(* IEC 61131-3 sources: codesys-framework/txt/application/ToDo/Hyperion, 15 files *)

(* ---- F_HyperionCreatePayloadString_1.pou.st ---- *)
FUNCTION F_HyperionCreatePayloadString_1 : ARRAY[0..63] OF BYTE
VAR_INPUT
	asEventPayload : ARRAY[1..10] OF STRING;
	iAmountPayload : INT;
END_VAR
VAR
	_sSeparator : STRING(1);
	_bySeparatorAsciiValue : BYTE;
	_byCharAsciiValue : BYTE;
	_iCounter : INT;
	_sPayloadPartString : STRING;
	_sPayloadString : STRING (cHYP_MAX_PAYLOADBYTESIZE);
	_iPayloadStringLength : INT;

	_abyPayloadByteArray : POINTER TO ARRAY [0 .. cHYP_MAX_PAYLOADBYTESIZE] OF BYTE;
	_abyPayloadByteArray_Return : ARRAY [0 .. cHYP_MAX_PAYLOADBYTESIZE] OF BYTE;
END_VAR

// --- BEGIN IMPLEMENTATION ---

// Init
_sPayloadString := '';
_sSeparator := ';';
_bySeparatorAsciiValue := 59;
// Check PayloadStrings
FOR _iCounter := 1 TO iAmountPayload BY 1 DO
	_sPayloadPartString := CONCAT(STR1 := asEventPayload[_iCounter], STR2 := _sSeparator);
	_sPayloadString := CONCAT(STR1 := _sPayloadString, STR2 := _sPayloadPartString);
END_FOR

// String to ByteArray
_iPayloadStringLength := LEN (STR := _sPayloadString);
_abyPayloadByteArray := ADR (_sPayloadString);

// Replace ';' with 0
FOR _iCounter := 0 TO cHYP_MAX_PAYLOADBYTESIZE BY 1 DO
	IF _iCounter < _iPayloadStringLength THEN
		_byCharAsciiValue := _abyPayloadByteArray^[_iCounter];
 		IF (_byCharAsciiValue <> _bySeparatorAsciiValue) THEN
			_abyPayloadByteArray_Return[_iCounter] := _byCharAsciiValue;
		ELSE
			_abyPayloadByteArray_Return[_iCounter] := 0;
		END_IF
	ELSE
		_abyPayloadByteArray_Return[_iCounter] := 0;
	END_IF
END_FOR

F_HyperionCreatePayloadString := _abyPayloadByteArray_Return;

(* ---- F_ParameterHandler_Bool.pou.st ---- *)
FUNCTION F_ParameterHandler_Bool : BOOL
VAR_INPUT
	eSubMachine 				: INT;
	w 							: WORD;
	eMode 						: E_ParameterMode;
	udiParameterId 				: UDINT;
	xExternalValidationFailed 	: BOOL := FALSE;
END_VAR
VAR_IN_OUT
	xValidationFailed 			: BOOL;
END_VAR
VAR_IN_OUT
	xHypValue 					: BOOL;
	xPLCValue 					: BOOL;
END_VAR
VAR
	_xParameterValid 			: BOOL;
	_rHypValue 					: REAL;
	_rPLCValue 					: REAL;
END_VAR

// --- BEGIN IMPLEMENTATION ---

IF (eMode = E_ParameterMode.Invalid) THEN
	xValidationFailed := TRUE;
	RETURN;
END_IF

IF xHypValue THEN
	_rHypValue := 1;
ELSE
	_rHypValue := 0;
END_IF

IF xPLCValue THEN
	_rPLCValue := 1;
ELSE
	_rPLCValue := 0;
END_IF

F_ParameterHandler_Real (
	eSubMachine := eSubMachine,
	w := w,
	eMode := eMode,
	udiParameterId := udiParameterId,
	xCanBeZero := TRUE,
	rLowLimit := 0,
	rUppLimit := 1,
	xValidationFailed := xValidationFailed,
	xExternalValidationFailed := xExternalValidationFailed,
	rHypValue := _rHypValue,
	rPLCValue := _rPLCValue);

xHypValue := _rHypValue = 1;
xPLCValue := _rPLCValue = 1;

(* ---- F_ParameterHandler_DInt.pou.st ---- *)
FUNCTION F_ParameterHandler_DInt : BOOL
VAR_INPUT
	eSubMachine 				: INT;
	w 							: WORD;
	eMode 						: E_ParameterMode;
	udiParameterId 				: UDINT;
	xCanBeZero 					: BOOL;
	diLowLimit 					: DINT;
	diUppLimit 					: DINT;
	xExternalValidationFailed 	: BOOL := FALSE;
END_VAR
VAR_IN_OUT
	xValidationFailed 			: BOOL;
	diHypValue 					: DINT;
	diPLCValue 					: DINT;
END_VAR
VAR
	_xParameterValid 			: BOOL;
	_rHypValue 					: REAL;
	_rPLCValue 					: REAL;
END_VAR

// --- BEGIN IMPLEMENTATION ---

IF eMode = E_ParameterMode.Invalid THEN
	xValidationFailed := TRUE;
	RETURN;
END_IF

_rHypValue := DINT_TO_REAL (diHypValue);
_rPLCValue := DINT_TO_REAL (diPLCValue);

F_ParameterHandler_Real (
	eSubMachine := eSubMachine,
	w := w,
	eMode := eMode,
	udiParameterId := udiParameterId,
	xCanBeZero := xCanBeZero,
	rLowLimit := DINT_TO_REAL (diLowLimit),
	rUppLimit := DINT_TO_REAL (diUppLimit),
	xValidationFailed := xValidationFailed,
	xExternalValidationFailed := xExternalValidationFailed,
	rHypValue := _rHypValue,
	rPLCValue := _rPLCValue);

diHypValue := REAL_TO_DINT (_rHypValue);
diPLCValue := REAL_TO_DINT (_rPLCValue);

(* ---- F_ParameterHandler_DWord.pou.st ---- *)
FUNCTION F_ParameterHandler_DWord : BOOL
VAR_INPUT
	eSubMachine 				: INT;
	w 							: WORD;
	eMode 						: E_ParameterMode;
	udiParameterId 				: UDINT;
	xCanBeZero 					: BOOL;
	dwLowLimit 					: DWORD;
	dwUppLimit 					: DWORD;
	xExternalValidationFailed 	: BOOL := FALSE;
END_VAR
VAR_IN_OUT
	xValidationFailed 			: BOOL;
	dwHypValue 					: DWORD;
	dwPLCValue 					: DWORD;
END_VAR
VAR
	_xParameterValid 			: BOOL;
	_rHypValue 					: REAL;
	_rPLCValue 					: REAL;
END_VAR

// --- BEGIN IMPLEMENTATION ---

IF eMode = E_ParameterMode.Invalid THEN
	xValidationFailed := TRUE;
	RETURN;
END_IF

_rHypValue := DWORD_TO_REAL (dwHypValue);
_rPLCValue := DWORD_TO_REAL (dwPLCValue);

F_ParameterHandler_Real (
	eSubMachine := eSubMachine,
	w := w,
	eMode := eMode,
	udiParameterId := udiParameterId,
	xCanBeZero := xCanBeZero,
	rLowLimit := DWORD_TO_REAL (dwLowLimit),
	rUppLimit := DWORD_TO_REAL (dwUppLimit),
	xValidationFailed := xValidationFailed,
	xExternalValidationFailed := xExternalValidationFailed,
	rHypValue := _rHypValue,
	rPLCValue := _rPLCValue);

dwHypValue := REAL_TO_DWORD (_rHypValue);
dwPLCValue := REAL_TO_DWORD (_rPLCValue);

(* ---- F_ParameterHandler_Int.pou.st ---- *)
FUNCTION F_ParameterHandler_Int : BOOL
VAR_INPUT
	eSubMachine 				: INT;
	w 							: WORD;
	eMode 						: E_ParameterMode;
	udiParameterId 				: UDINT;
	xCanBeZero 					: BOOL;
	iLowLimit 					: INT;
	iUppLimit 					: INT;
	xExternalValidationFailed 	: BOOL := FALSE;
END_VAR
VAR_IN_OUT
	xValidationFailed 			: BOOL;
	iHypValue 					: INT;
	iPLCValue 					: INT;
END_VAR
VAR
	_xParameterValid 			: BOOL;
	_rHypValue 					: REAL;
	_rPLCValue 					: REAL;
END_VAR

// --- BEGIN IMPLEMENTATION ---

IF eMode = E_ParameterMode.Invalid THEN
	xValidationFailed := TRUE;
	RETURN;
END_IF

_rHypValue := INT_TO_REAL (iHypValue);
_rPLCValue := INT_TO_REAL (iPLCValue);

F_ParameterHandler_Real (
	eSubMachine := eSubMachine,
	w := w,
	eMode := eMode,
	udiParameterId := udiParameterId,
	xCanBeZero := xCanBeZero,
	rLowLimit := INT_TO_REAL (iLowLimit),
	rUppLimit := INT_TO_REAL (iUppLimit),
	xValidationFailed := xValidationFailed,
	xExternalValidationFailed := xExternalValidationFailed,
	rHypValue := _rHypValue,
	rPLCValue := _rPLCValue);

iHypValue := REAL_TO_INT (_rHypValue);
iPLCValue := REAL_TO_INT (_rPLCValue);

(* ---- F_ParameterHandler_LReal.pou.st ---- *)
FUNCTION F_ParameterHandler_LReal : BOOL
VAR_INPUT
	eSubMachine 				: INT;
	w 							: WORD;
	eMode 						: E_ParameterMode;
	udiParameterId 				: UDINT;
	xCanBeZero 					: BOOL;
	lrLowLimit 					: LREAL;
	lrUppLimit 					: LREAL;
	xExternalValidationFailed 	: BOOL := FALSE;
END_VAR
VAR_IN_OUT
	xValidationFailed 			: BOOL;
	lrHypValue 					: LREAL;
	lrPLCValue 					: LREAL;
END_VAR
VAR
	_xParameterValid 			: BOOL;
END_VAR

// --- BEGIN IMPLEMENTATION ---

// Check
IF eMode = E_ParameterMode.Invalid THEN
	xValidationFailed := TRUE;
	RETURN;
END_IF

// Check HypValues
IF eMode = E_ParameterMode.CheckHyp THEN
	_xParameterValid := TRUE;
	IF NOT xCanBeZero AND lrHypValue = 0 THEN
		_xParameterValid := FALSE;
	ELSIF lrHypValue < lrLowLimit THEN
		_xParameterValid := FALSE;
	ELSIF lrHypValue > lrUppLimit THEN
		_xParameterValid := FALSE;
	ELSIF xExternalValidationFailed THEN
		_xParameterValid := FALSE;
	END_IF

	// !!!!! SET xParameterValidationFailed (Reset will be performed elsewhere)
	IF NOT _xParameterValid THEN
		xValidationFailed := TRUE;
	END_IF
END_IF

// Check PLCValues
IF eMode = E_ParameterMode.CheckPLC THEN
	_xParameterValid := TRUE;
	IF NOT xCanBeZero AND lrPLCValue = 0 THEN
		_xParameterValid := FALSE;
	ELSIF lrPLCValue < lrLowLimit THEN
		_xParameterValid := FALSE;
	ELSIF lrPLCValue > lrUppLimit THEN
		_xParameterValid := FALSE;
	ELSIF xExternalValidationFailed THEN
		_xParameterValid := FALSE;
	END_IF

	// !!!!! SET xParameterValidationFailed (Reset will be performed elsewhere)
	IF NOT _xParameterValid THEN
		xValidationFailed := TRUE;
	END_IF
END_IF

// Validate HyperionValues
IF eMode = E_ParameterMode.ValidateHyp OR eMode = E_ParameterMode.ValidateHypAndSavePLC THEN
	_xParameterValid := TRUE;
	IF NOT xCanBeZero AND lrHypValue = 0 THEN
		_xParameterValid := FALSE;
		// Insert message parametervalue is Zero
		F_Event_InsertMessage_ParameterChange (
			eSubMachine := eSubMachine,
			w := w,
			eValidationCode := E_ParameterValidationCode.Validation_Failed_IsZero,
			udiEventID := udiParameterId,
			rParameterValue_New := lrHypValue,
			rParameterValue_Previous := lrPLCValue,
			rParameterValue_MinimumValue := LREAL_TO_REAL(lrLowLimit),
			rParameterValue_MaximumValue := LREAL_TO_REAL(lrUppLimit));
	ELSIF lrHypValue < lrLowLimit THEN
		_xParameterValid := FALSE;
		//Insert message parametervalue < rValueLowerLimit
		F_Event_InsertMessage_ParameterChange (
			eSubMachine := eSubMachine,
			w := w,
			eValidationCode := E_ParameterValidationCode.Validation_Failed_BelowMinimum,
			udiEventID := udiParameterId,
			rParameterValue_New := lrHypValue,
			rParameterValue_Previous := lrPLCValue,
			rParameterValue_MinimumValue := LREAL_TO_REAL(lrLowLimit),
			rParameterValue_MaximumValue := LREAL_TO_REAL(lrUppLimit));
	ELSIF lrHypValue > lrUppLimit THEN
		_xParameterValid := FALSE;
		// Insert message parametervalue > rValueUpperLimit
		F_Event_InsertMessage_ParameterChange (
			eSubMachine := eSubMachine,
			w := w,
			eValidationCode := E_ParameterValidationCode.Validation_Failed_AboveMaximum,
			udiEventID := udiParameterId,
			rParameterValue_New := lrHypValue,
			rParameterValue_Previous := lrPLCValue,
			rParameterValue_MinimumValue := LREAL_TO_REAL(lrLowLimit),
			rParameterValue_MaximumValue := LREAL_TO_REAL(lrUppLimit));
	ELSIF xExternalValidationFailed THEN
		_xParameterValid := FALSE;
		// Insert message externalvalidationfailed
		F_Event_InsertMessage_ParameterChange (
			eSubMachine := eSubMachine,
			w := w,
			eValidationCode := E_ParameterValidationCode.Validation_Failed_External,
			udiEventID := udiParameterId,
			rParameterValue_New := lrHypValue,
			rParameterValue_Previous := lrPLCValue,
			rParameterValue_MinimumValue := LREAL_TO_REAL(lrLowLimit),
			rParameterValue_MaximumValue := LREAL_TO_REAL(lrUppLimit));
	END_IF

	// !!!!! SET xParameterValidationFailed (Reset will be performed elsewhere)
	IF NOT _xParameterValid THEN
		xValidationFailed := TRUE;
	END_IF
END_IF

// Save
IF eMode = E_ParameterMode.SavePLC OR (eMode = E_ParameterMode.ValidateHypAndSavePLC AND _xParameterValid) THEN
	IF lrPLCValue <> lrHypValue THEN
		F_Event_InsertMessage_ParameterChange (
			eSubMachine := eSubMachine,
			w := w,
			eValidationCode := E_ParameterValidationCode.Validation_Ok,
			udiEventID := udiParameterId,
			rParameterValue_New := lrHypValue,
			rParameterValue_Previous := lrPLCValue,
			rParameterValue_MinimumValue := LREAL_TO_REAL(lrLowLimit),
			rParameterValue_MaximumValue := LREAL_TO_REAL(lrUppLimit));
		lrPLCValue := lrHypValue;
	END_IF
END_IF

// Copy
IF eMode = E_ParameterMode.CopyPLCToHyp THEN
	lrHypValue := lrPLCValue;
END_IF

(* ---- F_ParameterHandler_Real.pou.st ---- *)
FUNCTION F_ParameterHandler_Real : BOOL
VAR_INPUT
	eSubMachine 				: INT;
	w 							: WORD;
	eMode 						: E_ParameterMode;
	udiParameterId 				: UDINT;
	xCanBeZero 					: BOOL;
	rLowLimit 					: REAL;
	rUppLimit 					: REAL;
	xExternalValidationFailed 	: BOOL := FALSE;
END_VAR
VAR_IN_OUT
	xValidationFailed 			: BOOL;
	rHypValue 					: REAL;
	rPLCValue 					: REAL;
END_VAR
VAR
	_xParameterValid 			: BOOL;
END_VAR

// --- BEGIN IMPLEMENTATION ---

// Check
IF eMode = E_ParameterMode.Invalid THEN
	xValidationFailed := TRUE;
	RETURN;
END_IF

// Check HypValues
IF eMode = E_ParameterMode.CheckHyp THEN
	_xParameterValid := TRUE;
	IF NOT xCanBeZero AND rHypValue = 0 THEN
		_xParameterValid := FALSE;
	ELSIF rHypValue < rLowLimit THEN
		_xParameterValid := FALSE;
	ELSIF rHypValue > rUppLimit THEN
		_xParameterValid := FALSE;
	ELSIF xExternalValidationFailed THEN
		_xParameterValid := FALSE;
	END_IF

	// !!!!! SET xParameterValidationFailed (Reset will be performed elsewhere)
	IF NOT _xParameterValid THEN
		xValidationFailed := TRUE;
	END_IF
END_IF

// Check PLCValues
IF eMode = E_ParameterMode.CheckPLC THEN
	_xParameterValid := TRUE;
	IF NOT xCanBeZero AND rPLCValue = 0 THEN
		_xParameterValid := FALSE;
	ELSIF rPLCValue < rLowLimit THEN
		_xParameterValid := FALSE;
	ELSIF rPLCValue > rUppLimit THEN
		_xParameterValid := FALSE;
	ELSIF xExternalValidationFailed THEN
		_xParameterValid := FALSE;
	END_IF

	// !!!!! SET xParameterValidationFailed (Reset will be performed elsewhere)
	IF NOT _xParameterValid THEN
		xValidationFailed := TRUE;
	END_IF
END_IF

// Validate HyperionValues
IF eMode = E_ParameterMode.ValidateHyp OR eMode = E_ParameterMode.ValidateHypAndSavePLC THEN
	_xParameterValid := TRUE;
	IF NOT xCanBeZero AND rHypValue = 0 THEN
		_xParameterValid := FALSE;
		// Insert message parametervalue is Zero
		F_Event_InsertMessage_ParameterChange (
			eSubMachine := eSubMachine,
			w := w,
			eValidationCode := E_ParameterValidationCode.Validation_Failed_IsZero,
			udiEventID := udiParameterId,
			rParameterValue_New := rHypValue,
			rParameterValue_Previous := rPLCValue,
			rParameterValue_MinimumValue := rLowLimit,
			rParameterValue_MaximumValue := rUppLimit);
	ELSIF rHypValue < rLowLimit THEN
		_xParameterValid := FALSE;
		//Insert message parametervalue < rValueLowerLimit
		F_Event_InsertMessage_ParameterChange (
			eSubMachine := eSubMachine,
			w := w,
			eValidationCode := E_ParameterValidationCode.Validation_Failed_BelowMinimum,
			udiEventID := udiParameterId,
			rParameterValue_New := rHypValue,
			rParameterValue_Previous := rPLCValue,
			rParameterValue_MinimumValue := rLowLimit,
			rParameterValue_MaximumValue := rUppLimit);
	ELSIF rHypValue > rUppLimit THEN
		_xParameterValid := FALSE;
		// Insert message parametervalue > rValueUpperLimit
		F_Event_InsertMessage_ParameterChange (
			eSubMachine := eSubMachine,
			w := w,
			eValidationCode := E_ParameterValidationCode.Validation_Failed_AboveMaximum,
			udiEventID := udiParameterId,
			rParameterValue_New := rHypValue,
			rParameterValue_Previous := rPLCValue,
			rParameterValue_MinimumValue := rLowLimit,
			rParameterValue_MaximumValue := rUppLimit);
	ELSIF xExternalValidationFailed THEN
		_xParameterValid := FALSE;
		// Insert message externalvalidationfailed
		F_Event_InsertMessage_ParameterChange (
			eSubMachine := eSubMachine,
			w := w,
			eValidationCode := E_ParameterValidationCode.Validation_Failed_External,
			udiEventID := udiParameterId,
			rParameterValue_New := rHypValue,
			rParameterValue_Previous := rPLCValue,
			rParameterValue_MinimumValue := rLowLimit,
			rParameterValue_MaximumValue := rUppLimit);
	END_IF

	// !!!!! SET xParameterValidationFailed (Reset will be performed elsewhere)
	IF NOT _xParameterValid THEN
		xValidationFailed := TRUE;
	END_IF
END_IF

// Save
IF eMode = E_ParameterMode.SavePLC OR (eMode = E_ParameterMode.ValidateHypAndSavePLC AND _xParameterValid) THEN
	IF rPLCValue <> rHypValue THEN
		F_Event_InsertMessage_ParameterChange (
			eSubMachine := eSubMachine,
			w := w,
			eValidationCode := E_ParameterValidationCode.Validation_Ok,
			udiEventID := udiParameterId,
			rParameterValue_New := rHypValue,
			rParameterValue_Previous := rPLCValue,
			rParameterValue_MinimumValue := rLowLimit,
			rParameterValue_MaximumValue := rUppLimit);
		rPLCValue := rHypValue;
	END_IF
END_IF

// Copy
IF eMode = E_ParameterMode.CopyPLCToHyp THEN
	rHypValue := rPLCValue;
END_IF

(* ---- F_ParameterHandler_String.pou.st ---- *)
FUNCTION F_ParameterHandler_String : BOOL
VAR_INPUT
	eSubMachine 				: INT;
	w 							: WORD;
	eMode 						: E_ParameterMode;
	udiParameterId 				: UDINT;
	xCanBeLengthZero 			: BOOL;
	iLowLengthLimit 			: INT;
	iUppLengthLimit 			: INT;
	xExternalValidationFailed 	: BOOL := FALSE;
END_VAR
VAR_IN_OUT
	xValidationFailed 			: BOOL;
	sHypValue 					: STRING;
	sPLCValue 					: STRING;
END_VAR
VAR
	_xParameterValid 			: BOOL;
	_sHypValue 					: STRING;
	_sPLCValue 					: STRING;
END_VAR

// --- BEGIN IMPLEMENTATION ---

_sHypValue := sHypValue;
_sPLCValue := sPLCValue;

// Check
IF (eMode = E_ParameterMode.Invalid) THEN
	xValidationFailed := TRUE;
	RETURN;
END_IF

// Check HypValues
IF (eMode = E_ParameterMode.CheckHyp) THEN
	_xParameterValid := TRUE;
	IF NOT xCanBeLengthZero AND (_sHypValue = '') THEN
		_xParameterValid := FALSE;
	ELSIF (LEN (_sHypValue) < iLowLengthLimit) THEN
		_xParameterValid := FALSE;
	ELSIF (LEN (_sHypValue) > iUppLengthLimit) THEN
		_xParameterValid := FALSE;
	ELSIF xExternalValidationFailed THEN
		_xParameterValid := FALSE;
	END_IF
	// !!!!!  SET xParameterValidationFailed (Reset will be performed elsewhere)
	IF (_xParameterValid = FALSE) THEN
		xValidationFailed := TRUE;
	END_IF
END_IF

//Check PLCValues
IF (eMode = E_ParameterMode.CheckPLC) THEN
	_xParameterValid := TRUE;
	IF (NOT xCanBeLengthZero AND (_sPLCValue = '')) THEN
		_xParameterValid := FALSE;
	ELSIF (LEN (_sPLCValue) < iLowLengthLimit) THEN
		_xParameterValid := FALSE;
	ELSIF (LEN (_sPLCValue) > iUppLengthLimit) THEN
		_xParameterValid := FALSE;
	ELSIF xExternalValidationFailed THEN
		_xParameterValid := FALSE;
	END_IF
	// !!!!!  SET xParameterValidationFailed (Reset will be performed elsewhere)
	IF NOT _xParameterValid THEN
		xValidationFailed := TRUE;
	END_IF
END_IF

// Validate HyperionValues
IF ((eMode = E_ParameterMode.ValidateHyp) OR (eMode = E_ParameterMode.ValidateHypAndSavePLC)) THEN
	_xParameterValid := TRUE;
	IF (NOT xCanBeLengthZero AND (_sHypValue = '')) THEN
		_xParameterValid := FALSE;
		// Insert message parametervalue is Zero
		F_Event_InsertMessage_StringParameterChange (
			eSubMachine := eSubMachine,
			w := w,
			udiEventID := udiParameterId,
			eValidationCode := E_ParameterValidationCode.Validation_Failed_IsZero,
			sParameterValue_Previous := _sPLCValue,
			sParameterValue_New := _sHypValue,
			iParameterValue_MinimumValue := iLowLengthLimit,
			iParameterValue_MaximumValue := iUppLengthLimit);
	ELSIF (LEN (_sHypValue) < iLowLengthLimit) THEN
		_xParameterValid := FALSE;
		// Insert message parametervalue < rValueLowerLimit
		F_Event_InsertMessage_StringParameterChange (
			eSubMachine := eSubMachine,
			w := w,
			udiEventID := udiParameterId,
			eValidationCode := E_ParameterValidationCode.Validation_Failed_BelowMinimum,
			sParameterValue_Previous := _sPLCValue,
			sParameterValue_New := _sHypValue,
			iParameterValue_MinimumValue := iLowLengthLimit,
			iParameterValue_MaximumValue := iUppLengthLimit);
	ELSIF (LEN (_sHypValue) > iUppLengthLimit) THEN
		_xParameterValid := FALSE;
		// Insert message parametervalue > rValueUpperLimit
		F_Event_InsertMessage_StringParameterChange (
			eSubMachine := eSubMachine,
			w := w,
			udiEventID := udiParameterId,
			eValidationCode := E_ParameterValidationCode.Validation_Failed_AboveMaximum,
			sParameterValue_Previous := _sPLCValue,
			sParameterValue_New := _sHypValue,
			iParameterValue_MinimumValue := iLowLengthLimit,
			iParameterValue_MaximumValue := iUppLengthLimit);
	ELSIF xExternalValidationFailed THEN
		_xParameterValid := FALSE;
		// Insert message external validatio nfailed
		F_Event_InsertMessage_StringParameterChange (
			eSubMachine := eSubMachine,
			w := w,
			udiEventID := udiParameterId,
			eValidationCode := E_ParameterValidationCode.Validation_Failed_External,
			sParameterValue_Previous := _sPLCValue,
			sParameterValue_New := _sHypValue,
			iParameterValue_MinimumValue := iLowLengthLimit,
			iParameterValue_MaximumValue := iUppLengthLimit);
	END_IF
	// !!!!!  SET xParameterValidationFailed (Reset will be performed elsewhere)
	IF NOT _xParameterValid THEN
		xValidationFailed := TRUE;
	END_IF
END_IF

// Save
IF ((eMode = E_ParameterMode.SavePLC) OR ((eMode = E_ParameterMode.ValidateHypAndSavePLC) AND _xParameterValid)) THEN
	IF (_sPLCValue <> _sHypValue) THEN
		F_Event_InsertMessage_StringParameterChange (
			eSubMachine := eSubMachine,
			w :=w,
			udiEventID := udiParameterId,
			eValidationCode := E_ParameterValidationCode.Validation_Ok,
			sParameterValue_Previous := _sPLCValue,
			sParameterValue_New := _sHypValue,
			iParameterValue_MinimumValue := iLowLengthLimit,
			iParameterValue_MaximumValue := iUppLengthLimit);
		_sPLCValue := _sHypValue;
	END_IF
END_IF

// Copy
IF (eMode = E_ParameterMode.CopyPLCToHyp) THEN
	_sHypValue := _sPLCValue;
END_IF

sHypValue := _sHypValue;
sPLCValue := _sPLCValue;

(* ---- F_ParameterHandler_UDInt.pou.st ---- *)
FUNCTION F_ParameterHandler_UDInt : BOOL
VAR_INPUT
	eSubMachine 				: INT;
	w 							: WORD;
	eMode 						: E_ParameterMode;
	udiParameterId	 			: UDINT;
	xCanBeZero 					: BOOL;
	udiLowLimit 				: UDINT;
	udiUppLimit 				: UDINT;
	xExternalValidationFailed 	: BOOL := FALSE;
END_VAR
VAR_IN_OUT
	xValidationFailed 			: BOOL;
	udiHypValue 				: UDINT;
	udiPLCValue 				: UDINT;
END_VAR
VAR
	_xParameterValid 			: BOOL;
	_rHypValue 					: REAL;
	_rPLCValue 					: REAL;
END_VAR

// --- BEGIN IMPLEMENTATION ---

IF eMode = E_ParameterMode.Invalid THEN
	xValidationFailed := TRUE;
	RETURN;
END_IF

_rHypValue := UDINT_TO_REAL (udiHypValue);
_rPLCValue := UDINT_TO_REAL (udiPLCValue);

F_ParameterHandler_Real (
	eSubMachine := eSubMachine,
	w := w,
	eMode := eMode,
	udiParameterId := udiParameterId,
	xCanBeZero := xCanBeZero,
	rLowLimit := UDINT_TO_REAL (udiLowLimit),
	rUppLimit := UDINT_TO_REAL (udiUppLimit),
	xValidationFailed := xValidationFailed,
	xExternalValidationFailed := xExternalValidationFailed,
	rHypValue := _rHypValue,
	rPLCValue := _rPLCValue);

udiHypValue := REAL_TO_UDINT (_rHypValue);
udiPLCValue := REAL_TO_UDINT (_rPLCValue);

(* ---- F_ParameterHandler_UInt.pou.st ---- *)
FUNCTION F_ParameterHandler_UInt : BOOL
VAR_INPUT
	eSubMachine 				: INT;
	w 							: WORD;
	eMode 						: E_ParameterMode;
	udiParameterId 				: UDINT;
	xCanBeZero 					: BOOL;
	uiLowLimit 					: UINT;
	uiUppLimit 					: UINT;
	xExternalValidationFailed 	: BOOL := FALSE;
END_VAR
VAR_IN_OUT
	xValidationFailed 			: BOOL;
	uiHypValue 					: UINT;
	uiPLCValue 					: UINT;
END_VAR
VAR
	_xParameterValid 			: BOOL;
	_rHypValue 					: REAL;
	_rPLCValue 					: REAL;
END_VAR

// --- BEGIN IMPLEMENTATION ---

IF eMode = E_ParameterMode.Invalid THEN
	xValidationFailed := TRUE;
	RETURN;
END_IF

_rHypValue := UINT_TO_REAL (uiHypValue);
_rPLCValue := UINT_TO_REAL (uiPLCValue);

F_ParameterHandler_Real (
	eSubMachine := eSubMachine,
	w := w,
	eMode := eMode,
	udiParameterId := udiParameterId,
	xCanBeZero := xCanBeZero,
	rLowLimit := UINT_TO_REAL (uiLowLimit),
	rUppLimit := UINT_TO_REAL (uiUppLimit),
	xValidationFailed := xValidationFailed,
	xExternalValidationFailed := xExternalValidationFailed,
	rHypValue := _rHypValue,
	rPLCValue := _rPLCValue);

uiHypValue := REAL_TO_UINT (_rHypValue);
uiPLCValue := REAL_TO_UINT (_rPLCValue);

(* ---- F_ParameterHandler_Word.pou.st ---- *)
FUNCTION F_ParameterHandler_Word : BOOL
VAR_INPUT
	eSubMachine 				: INT;
	w 							: WORD;
	eMode 						: E_ParameterMode;
	udiParameterId 				: UDINT;
	xCanBeZero 					: BOOL;
	wLowLimit 					: WORD;
	wUppLimit 					: WORD;
	xExternalValidationFailed 	: BOOL := FALSE;
END_VAR
VAR_IN_OUT
	xValidationFailed 			: BOOL;
	wHypValue 					: WORD;
	wPLCValue 					: WORD;
END_VAR
VAR
	_xParameterValid 			: BOOL;
	_rHypValue 					: REAL;
	_rPLCValue 					: REAL;
END_VAR

// --- BEGIN IMPLEMENTATION ---

IF eMode = E_ParameterMode.Invalid THEN
	xValidationFailed := TRUE;
	RETURN;
END_IF

_rHypValue := WORD_TO_REAL (wHypValue);
_rPLCValue := WORD_TO_REAL (wPLCValue);

F_ParameterHandler_Real (
	eSubMachine := eSubMachine,
	w := w,
	eMode := eMode,
	udiParameterId := udiParameterId,
	xCanBeZero := xCanBeZero,
	rLowLimit := WORD_TO_REAL (wLowLimit),
	rUppLimit := WORD_TO_REAL (wUppLimit),
	xValidationFailed := xValidationFailed,
	xExternalValidationFailed := xExternalValidationFailed,
	rHypValue := _rHypValue,
	rPLCValue := _rPLCValue);

wHypValue := REAL_TO_WORD (_rHypValue);
wPLCValue := REAL_TO_WORD (_rPLCValue);

(* ---- FB_Bistable_OrionButtonWithExternalEnable.pou.st ---- *)
FUNCTION_BLOCK FB_Bistable_OrionButtonWithExternalEnable
VAR_INPUT
	eSubMachine 			: INT;
	w 						: WORD;
	iIdNr 					: INT;
	udiSwitchOnEventID 		: UDINT;
	udiSwitchOffEventID 	: UDINT;
	udiDisabledEventID 		: UDINT;
	xButtonEnabled 			: BOOL;
END_VAR
VAR_IN_OUT
	udiButton 				: UDINT;
	xResetButton 			: BOOL;
END_VAR
VAR_OUTPUT
	xButtonPressed 			: BOOL;
END_VAR
VAR
END_VAR

// --- BEGIN IMPLEMENTATION ---

IF udiButton = 1 AND NOT xButtonPressed AND xButtonEnabled THEN
	F_Event_InsertMessage(eSubMachine := eSubMachine,w:=w, iComponentId := iIdNr, udiEventID := udiSwitchOnEventID, eEventLevel := E_EventLevels.EventIsInformational);
	xButtonPressed := TRUE;
	udiButton := 2;
END_IF

IF udiButton = 1 AND xButtonPressed THEN
	F_Event_InsertMessage(eSubMachine := eSubMachine,w:=w, iComponentId := iIdNr, udiEventID := udiSwitchOffEventID, eEventLevel := E_EventLevels.EventIsInformational);
	xButtonPressed := FALSE;
	udiButton := 0;
END_IF

IF udiButton = 1 AND NOT xButtonEnabled THEN
	F_Event_InsertMessage(eSubMachine := eSubMachine,w:=w, iComponentId := iIdNr, udiEventID := udiDisabledEventID, eEventLevel := E_EventLevels.EventIsInformational);
	xButtonPressed := FALSE;
	udiButton := 0;
END_IF

IF xResetButton THEN
	xButtonPressed := FALSE;
	xResetButton := FALSE;
	udiButton := 0;
END_IF

(* ---- FB_Bistable_OrionButtonWithExternalReset.pou.st ---- *)
FUNCTION_BLOCK FB_Bistable_OrionButtonWithExternalReset
VAR_INPUT
	eSubMachine 	: INT;
	w 				: WORD;
	iIdNr 			: INT;
	udiParameterId 	: UDINT;
END_VAR
VAR_IN_OUT
	udiButton 		: UDINT;
	xExternalReset 	: BOOL;
END_VAR
VAR_OUTPUT
	xButtonPressed 	: BOOL;
END_VAR
VAR
END_VAR

// --- BEGIN IMPLEMENTATION ---

//When button in Orion is clicked we receive value 1 on parameter udiButton
//If we write value 2 to parameter udiButton the button has a pressed appearance in Orion

IF udiButton = 1 AND NOT xButtonPressed THEN
	F_Event_InsertMessageString(eSubMachine := eSubMachine,w:=w, udiEventID := udiParameterId, eEventLevel := E_EventLevels.EventIsInformational, sMessageString1 := '1', sMessageString2 := '');
	xButtonPressed := TRUE;
	udiButton := 2;
END_IF

IF udiButton = 1 AND xButtonPressed THEN
	F_Event_InsertMessageString(eSubMachine := eSubMachine,w:=w, udiEventID := udiParameterId, eEventLevel := E_EventLevels.EventIsInformational, sMessageString1 := '0', sMessageString2 := '');
	xButtonPressed := FALSE;
	udiButton := 0;
END_IF

IF xExternalReset THEN
	xButtonPressed := FALSE;
	xExternalReset := FALSE;
	udiButton := 0;
END_IF

(* ---- FB_Monostable_OrionButton.pou.st ---- *)
FUNCTION_BLOCK FB_Monostable_OrionButton
VAR_INPUT
	eSubMachine 	: INT;
	w 				: WORD;
	iIdNr 			: INT;
	udiParameterId 	: UDINT;
END_VAR
VAR_IN_OUT
	udiButton 		: UDINT;
	xResetButton 	: BOOL;
END_VAR
VAR_OUTPUT
	xButtonPressed 	: BOOL;
END_VAR
VAR
END_VAR

// --- BEGIN IMPLEMENTATION ---

IF udiButton = 1 THEN
	xButtonPressed := TRUE;
	udiButton := 0;
	F_Event_InsertMessage(eSubMachine := eSubMachine,w:=w, iComponentId := iIdNr, udiEventID := udiParameterId, eEventLevel := E_EventLevels.EventIsInformational);
END_IF

IF xResetButton THEN
	xButtonPressed := FALSE;
	xResetButton := FALSE;
END_IF

(* ---- FB_Monostable_OrionButtonWithExternalEnable.pou.st ---- *)
FUNCTION_BLOCK FB_Monostable_OrionButtonWithExternalEnable
VAR_INPUT
	eSubMachine 		: INT;
	w 					: WORD;
	iIdNr 				: INT;
	udiSwitchOnEventID 	: UDINT;
	udiDisabledEventID 	: UDINT;
	xButtonEnabled 		: BOOL;
END_VAR
VAR_IN_OUT
	udiButton 			: UDINT;
	xResetButton 		: BOOL;
END_VAR
VAR_OUTPUT
	xButtonPressed 		: BOOL;
END_VAR
VAR
END_VAR

// --- BEGIN IMPLEMENTATION ---

IF udiButton = 1 AND xButtonEnabled THEN
	F_Event_InsertMessage(eSubMachine := eSubMachine,w:=w, iComponentId := iIdNr, udiEventID := udiSwitchOnEventID, eEventLevel := E_EventLevels.EventIsInformational);
	xButtonPressed := TRUE;
	udiButton := 0;
END_IF

IF udiButton = 1 AND NOT xButtonEnabled THEN
	F_Event_InsertMessage(eSubMachine := eSubMachine,w:=w, iComponentId := iIdNr, udiEventID := udiDisabledEventID, eEventLevel := E_EventLevels.EventIsInformational);
	xButtonPressed := FALSE;
	udiButton := 0;
END_IF

IF xResetButton THEN
	xButtonPressed := FALSE;
	xResetButton := FALSE;
	udiButton := 0;
END_IF
